FUNCTION F_SpindlePDSXLA170ClutchStatus : ET_SpindleClutchStatus
(*

The function used to get clutch status.

Constructor: 		Patryk Panylo
Company:		E. Riexinger GmbH
Date:			18.05.2018
Version:			1.00

Date:			Revision:		Who:				Comment
dd.mm.yyyy		x.xx			Initials			comment

*)
VAR_INPUT
	(* Input variables / Eingang Variablen *)
	stClutchStatus					:ST_SpindlePDSXLA170ClutchStatus; (* Clutch status  *)
END_VAR
VAR
	(* Variables *)

END_VAR


IF stClutchStatus.bRotatingS1 AND (stClutchStatus.bToolNotClampedS2 OR NOT stClutchStatus.bToolPresentS3 OR NOT stClutchStatus.bClutchInBaseS4)			(* Clutch rotating and not closed *)
THEN
	F_SpindlePDSXLA170ClutchStatus := ET_SpindleClutchStatus_RotatingNoClosed;

ELSIF NOT stClutchStatus.bToolNotClampedS2 AND NOT stClutchStatus.bToolPresentS3 AND stClutchStatus.bClutchInBaseS4			(* Clutch is closed without tool *)
THEN
	F_SpindlePDSXLA170ClutchStatus := ET_SpindleClutchStatus_ClosedWithoutTool;

ELSIF NOT stClutchStatus.bToolNotClampedS2 AND stClutchStatus.bToolPresentS3 AND stClutchStatus.bClutchInBaseS4				(* Clutch is closed with tool *)
THEN
	F_SpindlePDSXLA170ClutchStatus := ET_SpindleClutchStatus_ClosedWithTool;

ELSIF stClutchStatus.bToolNotClampedS2 AND NOT stClutchStatus.bToolPresentS3 AND NOT stClutchStatus.bClutchInBaseS4		(* Clutch is opened *)
THEN
	F_SpindlePDSXLA170ClutchStatus := ET_SpindleClutchStatus_Opened;

ELSE
	F_SpindlePDSXLA170ClutchStatus := ET_SpindleClutchStatus_NoDefined;
END_IF

END_FUNCTION

(* stored: Version 1.1.0.1, ProductVersion 3.1.4024.15
   POU F_SpindlePDSXLA170ClutchStatus: Id {a68537f7-012a-47b5-979a-24c748bdd043}, SpecialFunc None *)
